(* IEC 61131-3 sources: OpenPlc_Lezioni/contatore/build, 2 files *)

(* ---- plc.st ---- *)
TYPE
  LOGLEVEL : (CRITICAL, WARNING, INFO, DEBUG) := INFO;
END_TYPE

FUNCTION_BLOCK LOGGER
  VAR_INPUT
    TRIG : BOOL;
    MSG : STRING;
    LEVEL : LOGLEVEL := INFO;
  END_VAR
  VAR
    TRIG0 : BOOL;
  END_VAR

  IF TRIG AND NOT TRIG0 THEN
  {{
   LogMessage(GetFbVar(LEVEL),(char*)GetFbVar(MSG, .body),GetFbVar(MSG, .len));
  }}
  END_IF;
  TRIG0:=TRIG;
END_FUNCTION_BLOCK

PROGRAM program0
  VAR
    CTU0 : CTU;
  END_VAR
  VAR
    BT1 : BOOL;
    BT2 : BOOL;
    Led : BOOL;
  END_VAR
  VAR
    PV : INT := 5;
    R_TRIG1 : R_TRIG;
  END_VAR

  R_TRIG1(CLK := BT1);
  CTU0(CU := R_TRIG1.Q, R := BT2, PV := PV);
  Led := CTU0.Q;
END_PROGRAM

CONFIGURATION Config0

  RESOURCE Res0 ON PLC
    TASK task0(INTERVAL := T#20ms,PRIORITY := 0);
    PROGRAM instance0 WITH task0 : program0;
  END_RESOURCE
END_CONFIGURATION

(* ---- generated_plc.st ---- *)
PROGRAM program0
  VAR
    CTU0 : CTU;
  END_VAR
  VAR
    BT1 AT %IX100.0 : BOOL;
    BT2 AT %IX100.1 : BOOL;
    Led AT %QX100.0 : BOOL;
  END_VAR
  VAR
    PV : INT := 5;
    R_TRIG1 : R_TRIG;
  END_VAR

  R_TRIG1(CLK := BT1);
  CTU0(CU := R_TRIG1.Q, R := BT2, PV := PV);
  Led := CTU0.Q;
END_PROGRAM

CONFIGURATION Config0

  RESOURCE Res0 ON PLC
    TASK task0(INTERVAL := T#20ms,PRIORITY := 0);
    PROGRAM instance0 WITH task0 : program0;
  END_RESOURCE
END_CONFIGURATION
